(*
SPDX-FileCopyrightText: c 2026 Oleksandr Tiutyk <trofimich@gmail.com>
SPDX-License-Identifier: MIT
License: https://opensource.org/license/mit
*)

(*!
<summary>Checks positional removal and compaction of survivors.</summary>
<description>
Borrows a group-owned list reserved for this case. Use from one task at a stable address.
Teardown clears the list before publication.
</description>
*)

{attribute 'no_assign'}
{attribute 'no_explicit_call' := 'do not call this function block directly'}
FUNCTION_BLOCK ListRemoveAtTest EXTENDS TOF_Testing.SingleCycleTest
VAR_STAT
	{attribute 'hide'}
	_ClassName : STRING := __POUNAME();
END_VAR
VAR
	_List : TOF_Collections.IList;
END_VAR

(*!
<summary>Clears the fixture before the runner publishes the result.</summary>
<description>
Also runs after an unexpected exception interrupts the case.
</description>
*)
METHOD PROTECTED AfterTest
_List.Clear();
END_METHOD

//! <summary>Borrows the concrete class name. Callers must not modify it.</summary>
{attribute 'monitoring' := 'call'}
PROPERTY ClassName : REFERENCE TO STRING
GET
ClassName REF= _ClassName;
END_GET
END_PROPERTY

(*!
<summary>Checks positional removal and compaction of survivors.</summary>
*)
METHOD PROTECTED ExecuteTest
VAR
	values : ARRAY [0..5] OF STRING := ['String0', 'String1', 'String2', 'String3', 'String4', 'String5'];
	expected : ARRAY [0..4] OF STRING := ['String0', 'String1', 'String2', 'String4', 'String5'];
	i : DINT;
END_VAR
_List.AppendCopy(value := values[0]);
_List.AppendCopy(value := values[1]);
_List.AppendCopy(value := values[2]);
_List.AppendCopy(value := values[3]);
_List.AppendCopy(value := values[4]);
_List.AppendCopy(value := values[5]);

_List.RemoveAt(index := 3);

Assert.ThatDInt(
	actual := _List.Length,
	message := "Unexpected sequence after RemoveAt length"
).ToBe(expected := DINT#5);

FOR i := 0 TO 4 DO
	Assert.ThatString(
		actual := _List.Get(index := i).AsString255(),
		message := TOF_Core.WideStrings.Concat255("Unexpected sequence after RemoveAt at index ", TO_WSTRING(i))
	).ToBe(expected := expected[i]);
END_FOR
END_METHOD

(*!
<summary>Binds the list fixture for this case.</summary>
<description>
Stores a borrowed interface without invoking the fixture. The owning group keeps it alive and
reserves it for this case. TestElement initializes the name and parent.
</description>
<param name="name">Display name of this case.</param>
<param name="parent">Group that owns this case.</param>
<param name="list">Required live list reserved for this case.</param>
*)
METHOD FB_init : BOOL
VAR_INPUT
	bInitRetains: BOOL; // TRUE: the retain variables are initialized (reset warm / reset cold)
	bInCopyCode: BOOL; // TRUE: the instance will be copied to the copy code afterward (online change)
	name : WSTRING;
	parent : TOF_Testing.ITestElement;
	list : TOF_Collections.IList;
END_VAR
_List := list;
FB_init := TRUE;
END_METHOD

//! <summary>Borrows the compiler-initialized namespace name. Callers must not modify it.</summary>
{attribute 'monitoring' := 'call'}
PROPERTY NamespaceName : REFERENCE TO STRING
GET
NamespaceName REF= CurrentNamespace.Name;
END_GET
END_PROPERTY

//! <summary>Reports the concrete instance size in bytes.</summary>
{attribute 'monitoring' := 'call'}
PROPERTY SelfSize : ULINT
GET
SelfSize := XSIZEOF(THIS^);
END_GET
END_PROPERTY

END_FUNCTION_BLOCK

(* stored: Version 1.1.0.1, ProductVersion 3.1.4026.21
   POU ListRemoveAtTest: Id {a980d7c8-9f1e-4c57-94f4-9befde57da98}, SpecialFunc None
   Method AfterTest: Id {9ebbf083-18ce-4edc-99fe-71145ab07713}
   Property ClassName: Id {43d7cc80-0362-4f7d-a3ee-6ba85a9018b4}
   Get Get: Id {7fcb6fb6-cfa1-4e42-9207-65991c06d8f2}
   Method ExecuteTest: Id {a341f02a-9199-429b-9a92-2d1b0d147969}
   Method FB_init: Id {e8220f73-9338-4400-849b-ca52d3870c4b}
   Property NamespaceName: Id {b22c5728-33b9-454b-9774-98d4e3b96881}
   Get Get: Id {ed080213-16ad-4408-967d-b44a5ee14c66}
   Property SelfSize: Id {b8ca8269-fa58-44bd-af12-e30b5ad75e82}
   Get Get: Id {ade3d7da-2235-4328-992f-130312293275} *)
